VAR_GLOBAL CONSTANT
	mF_Mpc_degrees: DINT := 3;
	mF_Mpc_voff: LREAL := 0.0;
	mF_Mpc_yoff: LREAL := 0.0;
	mF_Mpc_RYscale: LREAL := 1.0;
	mF_Mpc_RMDscale: LREAL := 1.0;
	SS_INITIALIZE: SINT := 0;
	SS_STEP: SINT := 1;
END_VAR

(* stored: Version 1.1.0.1, ProductVersion 3.1.4024.9
   GVL GVL_1845925446: Id {d745f2f0-fda4-499d-a61d-8e2e5ff36590} *)
